Fanuc KAREL source: ko00073.KL

-- PROVISIONAL review KL for V1013-1; original PC SHA256 7bd3bd1e7e3213d103b52da7a770f1ee2493618d26b9ae1cc33cf5946ab67827
-- Incomplete behavior may be omitted. Consult companion uncertainty JSON. Do not deploy.
PROGRAM KO00073
%NOLOCKGROUP
BEGIN
  -- UNRESOLVED_PC offsets 5-12; opcodes 9D,23
  -- UNRESOLVED_PC offsets 17-66; opcodes 27,22,1C,27,49,7E,AD,22,31,7E,4A
  -- UNRESOLVED_PC offsets 71-75; opcodes 7F
END KO00073
